// Mitsubishi GX Works2 project: 후입우선회로   PLC: Q02/Q02H

PROGRAM MAIN
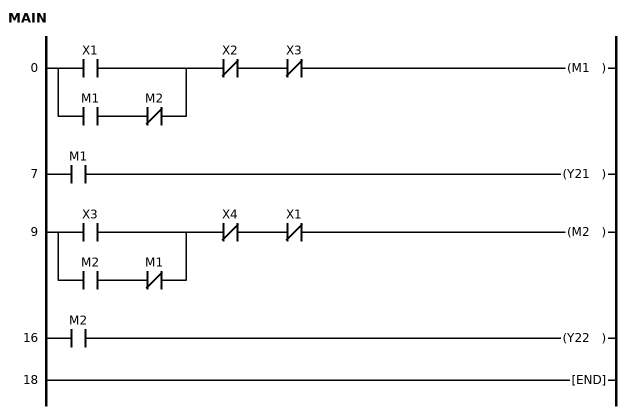
0     LD      X1
      LD      M1
      ANI     M2
      ORB
      ANI     X2
      ANI     X3
      OUT     M1
7     LD      M1
      OUT     Y21
9     LD      X3
      LD      M2
      ANI     M1
      ORB
      ANI     X4
      ANI     X1
      OUT     M2
16    LD      M2
      OUT     Y22
18    END
END_PROGRAM
